TYPE XtsModuleStatus :
STRUCT
	Module24Vdc: REAL;
	Module48Vdc: REAL;
	CurrentLive: LREAL;
	MaxCurrent: LREAL;
	ControlVdcOK : BOOL;
	MotorVdcOK : BOOL;
	ModuleInFault : BOOL;
	ModuleDriveState: Tc3_XTS_Utility.DriveState;
	ModuleCoEStatus: Tc3_XTS_Utility.CoeStatusInfo;
	ModuleEtherCATState: Tc3_XTS_Utility.EtherCatSlaveStateInfo;
	IsInfeed : BOOL;
END_STRUCT
END_TYPE

(* stored: Version 1.1.0.1
   DUT XtsModuleStatus: Id {7a4f3f27-a8bb-424a-97aa-0f14f7ad6bfd} *)
